(* ================================================================= *)
(*  FB_1012_ConveyorMotor                                             *)
(*  输送电机控制 - 方向互斥+慢速修饰+VFD故障检测                      *)
(*  版本: V9.0.0  日期: 2026-05-30                                    *)
(*  来源: SysLib/actuator/                                            *)
(*  规范: LSP-905-V1.0.2, LSP-904-V1.2.0, LSP-903-V1.0.0             *)
(*                                                                    *)
(*  V9.0.0变更 (Breaking Change):                                     *)
(*    - 重构: 移除VAR_IN_OUT ST_ConveyorMotor, 回归扁平接口           *)
(*    - 取消: 安全门信号(i_bSafetyDoorOk), 执行器不处理安全互锁       *)
(*    - 修正: 慢速改为方向修饰符, 必须与Fwd/Rev组合才生效             *)
(*    - 新增: 控制模式预留(i_iCtrlMode), 端子模式=0, 通讯模式=1       *)
(*    - 预留: 速度设定值(i_rSpeed), 通讯控制模式用                    *)
(* ================================================================= *)

FUNCTION_BLOCK FB_1012_ConveyorMotor

VAR_INPUT
    i_bFwdCmd       : BOOL;          // 正转命令
    i_bRevCmd       : BOOL;          // 反转命令
    i_bSlowCmd      : BOOL;          // 慢速命令(方向修饰符, 必须与Fwd/Rev组合)
    i_bVfdFault     : BOOL := FALSE; // 变频器故障输入
    i_iCtrlMode     : INT := 0;      // 控制模式: 0=端子控制, 1=通讯控制(预留)
    i_rSpeed        : REAL := 100.0; // 速度设定值(%, 通讯模式用, 端子模式无效)
END_VAR

VAR_OUTPUT
    q_bFwdOut       : BOOL;          // 正转输出(经互锁后)
    q_bRevOut       : BOOL;          // 反转输出(经互锁后)
    q_bSlowOut      : BOOL;          // 慢速输出(经互锁后)
    q_bRunning      : BOOL;          // 运行中
    q_bVfdAlarm     : BOOL;          // VFD报警
END_VAR

(* ==================== VFD故障检测 - 最高优先级 ==================== *)
IF i_bVfdFault THEN
    q_bVfdAlarm := TRUE;
    q_bFwdOut := FALSE;
    q_bRevOut := FALSE;
    q_bSlowOut := FALSE;
    q_bRunning := FALSE;
ELSE
    q_bVfdAlarm := FALSE;

    (* ==================== 方向命令仲裁 Fwd > Rev ==================== *)
    IF i_bFwdCmd THEN
        q_bFwdOut := TRUE;
        q_bRevOut := FALSE;
        q_bSlowOut := i_bSlowCmd;    // 慢速修饰正转
        q_bRunning := TRUE;
    ELSIF i_bRevCmd THEN
        q_bFwdOut := FALSE;
        q_bRevOut := TRUE;
        q_bSlowOut := i_bSlowCmd;    // 慢速修饰反转
        q_bRunning := TRUE;
    ELSE
        q_bFwdOut := FALSE;
        q_bRevOut := FALSE;
        q_bSlowOut := FALSE;         // 无方向命令时慢速无效
        q_bRunning := FALSE;
    END_IF;
END_IF;

END_FUNCTION_BLOCK
